Fanuc KAREL source: kt00039.KL

-- PROVISIONAL review KL for V940-1; original PC SHA256 e7853a1f9955603ec5d7f6a74c11b77c42e71b2e19a28e53fccd55a22ea1994b
-- Incomplete behavior may be omitted. Consult companion uncertainty JSON. Do not deploy.
PROGRAM KT00039
%NOLOCKGROUP
VAR
  I1 : INTEGER
  OUT : INTEGER
-- UNRESOLVED_DECL H2 type=002017
BEGIN
  -- V9_ZERO_TABLE_METADATA_HINT layout=0001; no indexed target words; source/name/runtime held
  -- UNRESOLVED_PC offsets 5-16; opcodes 2E,23
  -- UNRESOLVED_PC offsets 21-35; opcodes 2E,22,9D,33,B4
  -- UNRESOLVED_PC offsets 40-62; opcodes 21,22,9D,33,B3,53,23
  -- UNRESOLVED_PC offsets 67-71; opcodes 7F
END KT00039
